{attribute 'qualified_only'}
VAR_GLOBAL
	// Run/Stop Safety
	Run			AT%Q*:	BOOL;
	// Restart Safety
	Restart		AT%Q*:	BOOL;
	// Error Acknowledgement 
	ErrAck		AT%Q*:	BOOL;

END_VAR

(* stored: Version 1.1.0.1, ProductVersion 3.1.4024.13
   GVL GVL_Safety: Id {e2548b04-239f-4a51-958e-15ee3964bbc8} *)
